Universal Robots PolyScope program: Sub_Action_V2.urp

Program Sub_Action_V2 (installation=uLM011 MiR C1 BioRad directory=/programs/03 Sub Routines createdIn=5.16.0 lastSavedIn=5.16.0 robotSerialNumber=20245590045)
Calibrated DH parameters: a=[0.000135, -0.047884, -0.355309, -0.000204, 0.00003, 0]; d=[0.162633, 288.058298, -225.853183, -62.071663, 0.099761, 0.099601]; alpha=[1.569987, -0.001468, 0.002675, 1.570079, -1.570235, 0]; deltaTheta=[0, -1.458004, 8.179183, -0.437996, 0.000001, 0]
InitVariablesNode variables(variable(name=CMD_Abort, expression=False), variable(name=CMD_Clear, expression=False))
BeforeStart
  Script file /programs/04 Scripts/001 SCRIPT Errors and Warnings Deifnes V0.2.script
    | #*****************************************************
    | # customer          :   UK Essen
    | # project name      :   P1132
    | #****************************************************
    | # controller        :
    | # software          :
    | #****************************************************
    | # author            :   E.Petrichenko
    | # Copyright (c)     :   United Robotics Group Health and Food GmbH
    | #                       An der Riede 2
    | #                       28816 Stuhr
    | #                       Germany
    | #****************************************************
    | # description       :   centrifuge actions for the application
    | # version:      	:   0.1
    | # created           :   22.08.2024
    | # updated           :
    | #****************************************************
    | # modifications     :
    | #
    | # date              :
    | # name              :
    | # reason            :
    | #****************************************************
    | 
    | 
    | #################################### VARIABLES DEFINITIONS ###################################
    | 
    | ERROR_POSE_NOT_REACHABLE = 1002
    | ERROR_ROBOT_ARM_NOT_IN_HOME_POSE = 1006
    | ERROR_NO_OBJECT_TO_PICK = 1010
    | ERROR_NOT_DOCKED = 2003
    | ERROR_NOT_REACHABLE_TARGET = 2007
    | ERROR_CHARGING_NOT_STARTED = 2008
    | ERROR_AMR_WRONG_MODE = 2009
    | ERROR_UNKNOWN_POSE = 2010
    | ERROR_NO_LANDMARK = 3002
    | ERROR_WRONG_ORDER = 4002
    | ERROR_CENTRIFUGE_CONNECTION = 5001
    | ERROR_CENTRIFUGE_POWER = 5002
    | ERROR_CENTRIFUGE = 5003
    | ERROR_CENTRIFUGE_LID = 5004
    | ERROR_CANNOT_OPEN_HATCH = 5006
    | ERROR_CANNOT_CLOSE_HATCH = 5008
    | ERROR_CANNOT_ROTATE = 5010
    | ERROR_CANNOT_START = 5011
    | ERROR_WRONG_KEY_POSE = 5012
    | ERROR_MISSIING_CENTRACK = 5013
    | 
    | WARNING_POSE_NOT_REACHABLE = 1002
    | WARNING_BATTERY_LEVEL = 2002
    | WARNING_NOT_REACHABLE_TARGET = 2007
    | 
    | 
    | ERROR = struct(
    |     FLAG = False,
    |     ID = 0,
    |     MSG = "")
    | 
    | WARNING = struct(
    |     FLAG = False,
    |     ID = 0,
    |     MSG = "")
    | 
    | 
    | #################################### FUNCTIONS ###################################
    | 
    | def set_error(error_id):
    |     ERROR.ID = error_id
    |     if (ERROR.ID == 0):
    |         ERROR.FLAG = False
    |         ERROR.MSG = ""
    |     else:
    |         ERROR.FLAG = True
    |         if(ERROR.ID == ERROR_POSE_NOT_REACHABLE):
    |             ERROR.MSG = "Pose is not reachable"
    |         elif(ERROR.ID == ERROR_NO_OBJECT_TO_PICK):
    |             ERROR.MSG = "No object to pick"
    |         elif(ERROR.ID == ERROR_NO_LANDMARK):
    |             ERROR.MSG = "No landmark detected"
    |         elif(ERROR.ID == ERROR_ROBOT_ARM_NOT_IN_HOME_POSE):
    |             ERROR.MSG = "Robot arm cannot go to home pose"
    |         elif(ERROR.ID == ERROR_AMR_WRONG_MODE):
    |             ERROR.MSG = "AMR is in the wrong mode"
    |         elif(ERROR.ID == ERROR_NOT_DOCKED):
    |             ERROR.MSG = "Could not dock to the charger"
    |         elif(ERROR.ID == ERROR_NOT_REACHABLE_TARGET):
    |             ERROR.MSG = "Could not reach the target"
    |         elif(ERROR.ID == ERROR_CHARGING_NOT_STARTED):
    |             ERROR.MSG = "Could not start charging"
    |         elif(ERROR.ID == ERROR_UNKNOWN_POSE):
    |             ERROR.MSG = "Unknown navigation target"
    |         elif(ERROR.ID == ERROR_CANNOT_OPEN_HATCH):
    |             ERROR.MSG = "Centrifuge Cannot open the hatch"
    |         elif(ERROR.ID == ERROR_CENTRIFUGE_CONNECTION):
    |             ERROR.MSG = "Cannot reach centrifuge"
    |         elif (ERROR.ID == ERROR_CANNOT_CLOSE_HATCH):
    |             ERROR.MSG = "Centrifuge Cannot close the hatch"
    |         elif (ERROR.ID == ERROR_CANNOT_START):
    |             ERROR.MSG = "Centrifuge Cannot start"
    |         elif (ERROR.ID == ERROR_CANNOT_ROTATE):
    |             ERROR.MSG = "Centrifuge Cannot rotate the rotor"
    |         elif (ERROR.ID == ERROR_WRONG_ORDER):
    |             ERROR.MSG = "Wrong parameter was recieved"
    |         elif (ERROR.ID == ERROR_CENTRIFUGE):
    |             ERROR.MSG = "Centrifuge is in Error"
    |         elif (ERROR.ID == ERROR_WRONG_KEY_POSE):
    |             ERROR.MSG = "Key is in the wrong position"
    |         elif(ERROR.ID == ERROR_MISSIING_CENTRACK):
    |             ERROR.MSG = "Missing rack for centrifuge set"
    |         elif(ERROR.ID == ERROR_CENTRIFUGE_POWER):
    |             ERROR.MSG = "Centrifuge is turned off"
    |         elif(ERROR.ID == ERROR_CENTRIFUGE_LID):
    |             ERROR.MSG = "Lid of the centrifuge is opened"
    |         else:
    |             ERROR.MSG = "Unknown code"
    |         end
    |         textmsg("ERROR:",ERROR)
    |     end
    | end
    | 
    | def set_warning(warning_id):
    |     WARNING.ID = warning_id
    |     if (WARNING.ID == 0):
    |         WARNING.FLAG = False
    |         WARNING.MSG = ""
    |     else:
    |         WARNING.FLAG = True
    |         if(WARNING.ID == WARNING_POSE_NOT_REACHABLE):
    |             WARNING.MSG = "Pose is not reachable"
    |         elif(WARNING.ID == WARNING_BATTERY_LEVEL):
    |             WARNING.MSG = "Batery level dropped to a certain level"
    |         elif(WARNING.ID == WARNING_NOT_REACHABLE_TARGET):
    |             WARNING.MSG = "Not reachable location of AMR"
    |         else:
    |             WARNING.MSG = "Unknown code"
    |         end
    |         textmsg("WARNING:",WARNING)
    |     end
    | end
    | 
    | 
    | def reset_error():
    |   ERROR.ID = 0
    |   ERROR.FLAG = False
    |   ERROR.MSG = ""
    | end
    | 
    | 
    | def reset_warning():
    |     WARNING.ID = 0
    |     WARNING.FLAG = False
    |     WARNING.MSG = ""
    |   end
  Script file /programs/04 Scripts/SCRIPT Transitions V5.2.script
    | #*****************************************************
    | # customer          :   INTERNAL
    | # project name      :
    | #****************************************************
    | # controller        :   UR
    | # software          :   5.13
    | #****************************************************
    | # author            :   P. Koehnke
    | # Copyright (c)     :   United Robotics Group
    | #                       An der Riede 2
    | #                       28816 Stuhr
    | #                       Germany
    | #****************************************************
    | # description       :   transition between workareas
    | # version:      	:   1.2
    | # created           :   28.02.2024
    | # updated           :
    | #****************************************************
    | # modifications     :
    | #
    | # date              :
    | # name              :
    | # reason            :
    | #****************************************************
    | 
    | ######################### further development #########################
    | #   - that the robot can switch the configuration, if necessary
    | #   - introduction of structs
    | #######################################################################
    | 
    | ######################### to be adjusted #########################
    | local WORKAREA_1 = [-0.290,-0.560,-0.001, 0.290, 0.100, 1.000]    # workarea 1 (platform)
    | local WORKAREA_2 = [-1.000,-1.000,-1.000,-0.290, 0.100, 1.000]    # workarea 2 (front right)
    | local WORKAREA_3 = [-1.000, 0.100,-1.000, 0.000, 1.000, 1.000]    # workarea 3 (back right)
    | local WORKAREA_4 = [ 0.000, 0.100,-1.000, 1.000, 1.000, 1.000]    # workarea 4 (back left)
    | local WORKAREA_5 = [ 0.290,-1.000,-1.000, 1.000, 0.100, 1.000]    # workarea 5 (front left)
    | local WORKAREA_6 = [-0.290,-1.000,-1.000, 0.290,-0.560, 1.000]    # workarea 6 (front front)
    | local WORKAREA_7 = [0,0,0,0,0,0]    # reserved
    | local WORKAREA_8 = [0,0,0,0,0,0]    # reserved
    | local WORKAREA_9 = [0,0,0,0,0,0]    # reserved
    | local WORKAREA_10 = [0,0,0,0,0,0]   # reserved
    | 
    | local PSE_WA_1 = p[ 0.000,-0.400, 0.300, 0.000, 0.000, 0.000]
    | local PSE_WA_2 = p[-0.300,-0.300, 0.300, 0.000, 0.000, d2r(-90)]
    | local PSE_WA_3 = p[-0.300, 0.300, 0.300, 0.000, 0.000, d2r(-135)]
    | local PSE_WA_4 = p[ 0.300, 0.300, 0.300, 0.000, 0.000, d2r(135)]
    | local PSE_WA_5 = p[ 0.300,-0.300, 0.300, 0.000, 0.000, d2r(90)]
    | local PSE_WA_6 = p[ 0.000,-0.600, 0.300, 0.000, 0.000, 0.000]       # reserved
    | local PSE_WA_7 = p[ 0.000, 0.000, 0.000, 0.000, 0.000, 0.000]       # reserved
    | local PSE_WA_8 = p[ 0.000, 0.000, 0.000, 0.000, 0.000, 0.000]       # reserved
    | local PSE_WA_9 = p[ 0.000, 0.000, 0.000, 0.000, 0.000, 0.000]       # reserved
    | local PSE_WA_10 = p[ 0.000, 0.000, 0.000, 0.000, 0.000, 0.000]      # reserved
    | 
    | local JNT_STANDARD_C1 = [ 1.57,-1.57, 1.57,-1.57,-1.57,0]
    | local JNT_STANDARD_C2 = [-1.57,-1.57,-1.57,-1.57, 1.57,0]
    | local CLEARANCE_STANDARD = [-0.500,-0.900,-1.000, 0.500, 0.900, 1.000]  # desired free space around the base
    | local DISTANCE_TO_CLEARANCE = 0.300
    | local RADIUS_HELPER_POSES = 0.250
    | local RADIUS_TRANSITION_POSES = 0.400
    | local workareas = [WORKAREA_1, WORKAREA_2, WORKAREA_3, WORKAREA_4, WORKAREA_5, WORKAREA_6, WORKAREA_7, WORKAREA_8, WORKAREA_9, WORKAREA_10]
    | local poses = [PSE_WA_1, PSE_WA_2, PSE_WA_3, PSE_WA_4, PSE_WA_5, PSE_WA_6, PSE_WA_7, PSE_WA_8, PSE_WA_9, PSE_WA_10]
    | 
    | ######################### end of adjustment #########################
    | 
    | local pi = 3.14159265
    | local axis_config_current = 0
    | local axis_config_new = 0
    | local workarea_current = 0
    | local workarea_new = 0
    | local reverse_rotation = False
    | local yaw_locked =  0
    | local pose_start = struct(crt = p[0,0,0,0,0,0], jnt = [0,0,0,0,0,0], q = [0,0,0,0,0,0])
    | local pose_help = struct(crt = p[0,0,0,0,0,0], jnt = [0,0,0,0,0,0], q = [0,0,0,0,0,0])
    | local pose_target = struct(crt = p[0,0,0,0,0,0], jnt = [0,0,0,0,0,0], q = [0,0,0,0,0,0])
    | local pose = struct(crt = p[0,0,0,0,0,0], jnt = [0,0,0,0,0,0], q = [0,0,0,0,0,0])
    | 
    | def get_tool_free_pose(pose_ref=get_actual_tcp_pose(), dir=[0,0,0], move_in_base_frame=False):
    |     # get a recovery pose
    |     # dir is providing the direction and distance in X, Y and Z
    |     # if 'move_in_base_frame' is set, dir will be interpreted as absolute values for a movement in base frame
    | 
    |     local pose_target = pose_ref
    |     local i = 0
    | 
    |     if (move_in_base_frame):
    |         while (i<3):
    |             # move only,
    |             # if the demanded position is bigger than zero and the current position is below the demanded one or
    |             # if the demanded position is smaller than zero and the current position is above the demanded one
    |             if ((dir[i]>0 and pose_ref[i]<dir[i]) or (dir[i]<0 and pose_ref[i]>dir[i])):
    |                 pose_target[i] = dir[i]
    |             end
    |             i = i + 1
    |         end
    |     else:
    |         pose_target = pose_trans(pose_ref, p[dir[0], dir[1], dir[2], 0, 0, 0])
    |     end
    | 
    |     return pose_target
    | end
    | 
    | def check_workarea(reference_pose):
    |     # the actual TCP position is compared to predefined areas (cubic) to determine in which area the robot arm is
    |     # a workarea is defined as a list of coordinates, where the first 3 values are X, Y, and Z with the smallest values and
    |     # the next 3 values specify X, Y and Z for the biggest values
    | 
    |     local data_size = size(workareas)
    |     local i = 0
    |     local size_workarea = p[0,0,0,0,0,0]
    |     local pose_workarea = p[0,0,0,0,0,0]
    | 
    |     while (i < data_size[0]):
    |         pose_workarea = pose_trans(inv(p[workareas[i, 0], workareas[i, 1], workareas[i, 2], 0, 0, 0]), reference_pose)
    |         size_workarea = pose_sub(p[workareas[i, 3], workareas[i, 4], workareas[i, 5], 0, 0, 0], p[workareas[i, 0], workareas[i, 1], workareas[i, 2], 0, 0, 0])
    |         if  ((pose_workarea[0]>0 and pose_workarea[0]<size_workarea[0]) and
    |             (pose_workarea[1]>0 and pose_workarea[1]<size_workarea[1]) and
    |             (pose_workarea[2]>0 and pose_workarea[2]<size_workarea[2])):
    |             return i + 1
    |         end
    |         i = i + 1
    |     end
    |     return 0
    | end
    | 
    | def check_current_axis_config():
    |     # function determnines, if the arm is oriented in one or the other configuration.
    |     # it means, that the ellbow joint is flipped and so are the wrist joints.
    | 
    |     local jnt_current = get_actual_joint_positions()
    | 
    |     # ellbow has positiv angle
    |     if (jnt_current[2]> 0):
    |         return 1
    |     # ellbow has negativ angle
    |     elif (jnt_current[2]< 0):
    |         return 2
    |     # angle is 0
    |     else:
    |         return 0
    |     end
    | end
    | 
    | def switch_axis_config(axis_config):
    |     # function to switch betwwen the axis configuration 1 and 2.
    | 
    |     if (axis_config == 1):
    |         return 2
    |     elif (axis_config ==2):
    |         return 1
    |     end
    | end
    | 
    | def get_transition_pose(workarea, axis_config, closest=False, keep_xyz=[False, False, False]):
    |     # get the correspondig pose from the list of poses
    | 
    |     local jnt_current = get_actual_joint_positions()
    |     local pose_current = get_actual_tcp_pose()
    |     local i = 0
    | 
    |     pose.crt = poses[workarea-1]
    |     # if wanted, the pose will take the current position as desired x, y and z
    |     while (i < 3):
    |         if keep_xyz[i]:
    |             pose.crt[i] = pose_current[i]
    |         end
    |         i = i + 1
    |     end
    | 
    |     if (axis_config == 1):
    |         pose.q = JNT_STANDARD_C1
    |     elif (axis_config == 2):
    |         pose.q = JNT_STANDARD_C2
    |     end
    | 
    |     if closest:
    |         pose.q[0] = jnt_current[0]
    |     end
    | 
    |     if get_inverse_kin_has_solution(pose.crt, qnear=pose.q):
    |         pose.jnt = get_inverse_kin(pose.crt, qnear=pose.q)
    |     else:
    |         popup("no solution found for the transition pose", blocking= True)
    |     end
    | 
    |     return pose
    | end
    | 
    | def get_transition_pose_2(ref, radius, axis_config, closest=False):
    |     # get the correspondig pose from the list of poses
    | 
    |     local jnt_current = get_actual_joint_positions()
    |     local yaw_current = get_yaw_too_base(ref)
    | 
    |     #pose.crt = get_tool_free_pose(pose_ref=ref, dir=[0, 0, DISTANCE_TO_CLEARANCE], move_in_base_frame=True)
    | 
    |     if (axis_config == 1):
    |         pose.q = JNT_STANDARD_C1
    |     elif (axis_config == 2):
    |         pose.q = JNT_STANDARD_C2
    |     end
    | 
    |     if closest:
    |         pose.q[0] = jnt_current[0]
    |     end
    | 
    |     # get coordinates of the circle with the same angle as the given pose to the
    |     if ref == p[0,0,0,0,0,0]:
    |         pose.crt = PSE_WA_1
    |     else:
    |         pose.crt =
    |         p[radius * cos(yaw_current-pi/2),
    |         radius * sin(yaw_current-pi/2),
    |         DISTANCE_TO_CLEARANCE,
    |         0,
    |         0,
    |         yaw_current + get_locked_yaw()]
    |     end
    | 
    |     if get_inverse_kin_has_solution(pose.crt, qnear=pose.q):
    |         pose.jnt = get_inverse_kin(pose.crt, qnear=pose.q)
    |         #return pose
    |     else:
    |         popup("no solution found for the transition pose", blocking= True)
    |     end
    | 
    |     return pose
    | end
    | 
    | def get_rounded_mm(value):
    |     if (value < 0):
    |         return ceil(value*1000)
    |     elif (value >= 0):
    |         return floor(value*1000)
    |     end
    | end
    | 
    | def get_yaw_too_base(pose):
    |     # get the yaw relative to the base frame
    |     local pose_x_mm = 0
    |     local pose_y_mm = 0
    |     local yaw = 0
    | 
    |     pose_x_mm = get_rounded_mm(pose[0])
    |     pose_y_mm = get_rounded_mm(pose[1])
    | 
    |     if (pose_x_mm == 0 and pose_y_mm < 0):
    |         yaw = 0
    |     elif (pose_x_mm == 0 and pose_y_mm > 0):
    |         yaw = pi
    |     elif (pose_x_mm < 0 and pose_y_mm == 0):
    |         yaw = -pi/2
    |     elif (pose_x_mm > 0 and pose_y_mm == 0):
    |         yaw = pi/2
    |     else:
    |         yaw = atan2(pose[0], pose[1])
    |         if (-pi < yaw) and (yaw < 0):
    |             yaw = - yaw - pi
    |         elif (0 < yaw) and (yaw < pi):
    |             yaw = - yaw + pi
    |         else:
    |             yaw = pi
    |         end
    |     end
    |     return yaw
    | end
    | 
    | def get_helper_pose():
    |     # get the helper pose, as described
    | 
    |     local m_line = 0                    # slope of the line between base and circle point
    |     local n = 0                         # shift on the ordinate axis
    |     local m_normal = 0                  # slope of the normal of the line between base and circle point
    |     local x_p1 = 0                      # x coordinate of first circle point
    |     local x_p2 = 0                      # x coordinate of second circle point
    |     local y_p1 = 0                      # y coordinate of first circle point
    |     local y_p2 = 0                      # y coordinate of second circle point
    |     local jnt_help_1 = [0,0,0,0,0,0]
    |     local jnt_help_2 = [0,0,0,0,0,0]
    | 
    |     if (pose_start.crt != pose_target.crt):
    |         if (pose_start.crt[0] == pose_target.crt[0]):
    |             m_normal = 0
    |         elif (pose_start.crt[0] != pose_target.crt[0]):
    |             m_line = (pose_target.crt[1]-pose_start.crt[1])/(pose_target.crt[0]-pose_start.crt[0])    # calculation of the slope between start and target
    |             n = pose_start.crt[1] - m_line * pose_start.crt[0]
    |         end
    |         if (-0.00001 > m_line or m_line > 0.00001):
    |             m_normal = -1/m_line
    |         end
    | 
    |         # using p-q-formula for getting the crossing points
    |         x_p1 = sqrt(pow(RADIUS_HELPER_POSES, 2)/(pow(m_normal, 2)+1)) * -1
    |         x_p2 = sqrt(pow(RADIUS_HELPER_POSES, 2)/(pow(m_normal, 2)+1))
    |         y_p1 = m_normal * x_p1
    |         y_p2 = m_normal * x_p2
    |         pose.q = pose_start.jnt
    | 
    |         if (point_dist(pose_start.crt, p[x_p1, y_p1,0,0,0,0]) < point_dist(pose_start.crt, p[x_p2, y_p2,0,0,0,0])):
    |             if reverse_rotation:
    |                 pose_help.crt[0] = x_p2
    |                 pose_help.crt[1] = y_p2
    |                 pose.q = pose_target.jnt
    |             else:
    |                 pose_help.crt[0] = x_p1
    |                 pose_help.crt[1] = y_p1
    |                 pose.q = pose_start.jnt
    |             end
    |         elif (point_dist(pose_start.crt, p[x_p1, y_p1,0,0,0,0]) > point_dist(pose_start.crt, p[x_p2, y_p2,0,0,0,0])):
    |             if reverse_rotation:
    |                 pose_help.crt[0] = x_p1
    |                 pose_help.crt[1] = y_p1
    |                 pose.q = pose_target.jnt
    |             else:
    |                 pose_help.crt[0] = x_p2
    |                 pose_help.crt[1] = y_p2
    |                 pose.q = pose_start.jnt
    |             end
    |         elif (point_dist(pose_start.crt, p[x_p1, y_p1,0,0,0,0]) == point_dist(pose_start.crt, p[x_p2, y_p2,0,0,0,0])):
    |             jnt_help_1 = get_inverse_kin(p[x_p1, y_p1,pose_start.crt[2],pose_start.crt[3],pose_start.crt[4],pose_start.crt[5]], qnear=pose.q)
    |             jnt_help_2 = get_inverse_kin(p[x_p2, y_p2,pose_start.crt[2],pose_start.crt[3],pose_start.crt[4],pose_start.crt[5]], qnear=pose.q)
    |             if (pose_start.jnt[0]<jnt_help_1[0] and jnt_help_1[0]<pose_target.jnt[0]) or (pose_start.jnt[0]>jnt_help_1[0] and jnt_help_1[0]>pose_target.jnt[0]):
    |                 pose_help.crt[0] = x_p1
    |                 pose_help.crt[1] = y_p1
    |             elif (pose_start.jnt[0]<jnt_help_2[0] and jnt_help_2[0]<pose_target.jnt[0]) or (pose_start.jnt[0]>jnt_help_2[0] and jnt_help_2[0]>pose_target.jnt[0]):
    |                 pose_help.crt[0] = x_p2
    |                 pose_help.crt[1] = y_p2
    |             end
    |             pose.q = pose_start.jnt
    |         end
    | 
    |         pose_help.crt[2] = 0.5 * (pose_start.crt[2] + pose_target.crt[2])
    | 
    |         if ((pose_start.crt[1] < 0 and pose_target.crt[1] > 0) or (pose_start.crt[1] > 0 and pose_target.crt[1] < 0)):
    |             if get_inverse_kin_has_solution(pose.crt, qnear=pose.q):
    |                 pose.jnt = get_inverse_kin(pose.crt, qnear=pose.q)
    |             else:
    |                 popup("no solution found for the helper pose", blocking= True)
    |             end
    |         end
    |     end
    |     return pose
    | end
    | 
    | def adjust_transition_poses(pose_identifier):
    |     # adjust the orientation of the transition poses by determining the the current orientation
    | 
    |     local pose_current = get_actual_tcp_pose()
    |     local jnt_current = get_actual_joint_positions()
    |     local rpy_current = rotvec2rpy([pose_current[3],pose_current[4],pose_current[5]])
    |     local rotvec_new = [0,0,0]
    | 
    |     if (pose_identifier == "start"):
    |         pose.q = pose_start.jnt
    |         pose.crt = get_forward_kin(pose_start.jnt)
    |     elif (pose_identifier == "helper"):
    |         pose.q = pose_help.jnt
    |         pose.crt = get_forward_kin(pose_help.jnt)
    |     elif (pose_identifier == "target"):
    |         pose.q = pose_target.jnt
    |         pose.crt = get_forward_kin(pose_target.jnt)
    |     end
    | 
    |     rotvec_new = rpy2rotvec([rpy_current[0], rpy_current[1], get_yaw_too_base(pose.crt) + yaw_locked])
    |     pose.crt = p[pose.crt[0], pose.crt[1], pose.crt[2], rotvec_new[0], rotvec_new[1], rotvec_new[2]]
    | 
    |     pose.q[3] = jnt_current[3]
    |     pose.q[4] = jnt_current[4]
    |     pose.q[5] = jnt_current[5]
    |     if get_inverse_kin_has_solution(pose.crt, qnear=pose.q) and is_within_safety_limits(pose.crt):
    |         pose.jnt = get_inverse_kin(pose.crt, qnear=pose.q)
    |     else:
    |         popup(str_cat("no solution for ", pose_identifier), error=True, blocking=True)
    |     end
    |     return pose.jnt
    | end
    | 
    | def get_locked_yaw():
    |     local pose_current = get_actual_tcp_pose()
    |     local rpy_current = rotvec2rpy([pose_current[3],pose_current[4],pose_current[5]])
    |     local rotvec_new = rpy2rotvec([rpy_current[0], rpy_current[1], get_yaw_too_base(pose_current)])
    |     local pose_reference = p[pose_current[0], pose_current[1], pose_current[2], rotvec_new[0], rotvec_new[1], rotvec_new[2]]
    |     local pose_to_reference = pose_trans(pose_inv(pose_reference), get_actual_tcp_pose())
    |     yaw_locked = pose_to_reference[5]
    | 
    |     return yaw_locked
    | end
    | 
    | def do_transition(reference_pose=p[0,0,0,0,0,0], mode=2, keep_xyz=[False, False, False], keep_rxry=False, a=1.4, v=1.05, r=0.100):
    |     # the robot will evaluate the current and target workarea
    |     # after that, the robot will move between the workareas automatically.
    |     # parameters:
    |     # reference_pose:   a pose/frame were the robot should work next. If nothing is given, base frame will be used as target
    |     # keep_rxry:        if true, the robot will keep the orientation of the tool during the movement
    | 
    |     ################# checking #################
    |     axis_config_current = check_current_axis_config()           # 0: unknown, 1: config 1, 2: config 2
    |     workarea_current = check_workarea(get_actual_tcp_pose())    # between 0 and the amount of defined workareas
    |     workarea_new = check_workarea(reference_pose)               # between 0 and the amount of defined workareas
    |     if(workarea_current==workarea_new):
    |          return 0
    |     end
    |     if (workarea_current != 0 and workarea_new != 0):
    |         ################# get axisvalues #################
    |         # pose_start = get_transition_pose(workarea_current, axis_config_current, closest=not reverse_rotation, keep_xyz=keep_xyz)
    |         pose_start = get_transition_pose_2(get_actual_tcp_pose(), RADIUS_TRANSITION_POSES, axis_config_current, closest=not reverse_rotation)
    |         if (workarea_current == 3 and workarea_new == 4) or (workarea_current == 4 and workarea_new == 3):
    |             # pose_target = get_transition_pose(workarea_new, axis_config_current, closest=True)
    |             pose_target = get_transition_pose_2(reference_pose, RADIUS_TRANSITION_POSES, axis_config_current, closest=True)
    |             reverse_rotation = True
    |         else:
    |             pose_target = get_transition_pose_2(reference_pose, RADIUS_TRANSITION_POSES, axis_config_current, closest=(workarea_current == workarea_new))
    |             if reverse_rotation:
    |                 reverse_rotation = False
    |             end
    |         end
    |         # pose_help = get_helper_pose()
    |         global A_Start = pose_start.crt
    |         global A_Help = pose_help.crt
    |         global A_End = pose_target.crt
    | 
    | 
    |         ################# adjustments #################
    |         if (keep_rxry):
    |             get_locked_yaw()
    |             if (pose_start.jnt == pose_target.jnt):
    |                 pose_target.jnt = adjust_transition_poses("target")
    |                 pose_start.jnt = pose_target.jnt
    |             else:
    |                 pose_start.jnt = adjust_transition_poses("start")
    |                 pose_target.jnt = adjust_transition_poses("target")
    |             end
    |             if (pose_help.jnt != [0,0,0,0,0,0]):
    |                 pose_help.jnt = adjust_transition_poses("helper")
    |             end
    |         end
    | 
    |         global A_Start = pose_start.crt
    |         global A_Help = pose_help.crt
    |         global A_End = pose_target.crt
    | 
    |         ################# movements #################
    | 
    |         if point_dist(pose_start.crt, pose_target.crt) > 0.100:
    |             movej(pose_start.jnt, a=a, v=v, r=r)
    |         end
    |         # if (pose_help.jnt != [0,0,0,0,0,0]):
    |         #     movej(pose_help.jnt, a=a, v=v, r=r)
    |         # end
    |         movej(pose_target.jnt, a=a, v=v)
    |     else:
    |         # define error
    |     end
    | 
    |     ################# checking #################
    |     axis_config_current = check_current_axis_config()           # 0: unknown, 1: config 1, 2: config 2
    |     workarea_current = check_workarea(get_actual_tcp_pose())    # between 0 and the amount of defined workareas
    | end
  Script file /programs/04 Scripts/SCRIPT Utility V5.1.script
    | #*****************************************************
    | # customer          :   tbd
    | # project name      :   tbd
    | #****************************************************
    | # controller        :
    | # software          :
    | #****************************************************
    | # author            :   P. Koehnke (+49 1628859904; p.koehnke@unitedrobotics.group)
    | # Copyright (c)     :   United Robotics Group Health and Food GmbH
    | #                       An der Riede 2
    | #                       28816 Stuhr
    | #                       Germany
    | #****************************************************
    | # description       :   utility programs for the application
    | # version:      	:   3.1
    | # created           :   30.01.2023
    | # updated           :
    | #****************************************************
    | # modifications     :   get_tool_free_pose_2(), get_index_from_list()
    | #
    | # date              :   05.01.2024
    | # name              :   PK
    | # reason            :
    | #****************************************************
    | 
    | def found_in_matrix(data, req_id, req_idx):
    |     local id = -1
    |     local dimensions = size(data)
    |     local loop_dataset = 0
    | 
    |     while (id != req_id and loop_dataset < dimensions[0]):
    |         id = data[loop_dataset, 0]
    |         if (id == req_id):
    |             return data[loop_dataset, req_idx]
    |         else:
    |             loop_dataset = loop_dataset + 1
    |         end
    |     end
    | end
    | 
    | def found_in_list(value, list):
    |     local idx = 0
    | 
    |     while (idx < length(list)):
    |         if (value == list[idx]):
    |             return True
    |         end
    |         idx = idx + 1
    |     end
    |     return False
    | end
    | 
    | def get_index_from_list(list, value=-1):
    |     local idx = 0
    | 
    |     while (idx < length(list)):
    |         if (value == -1):
    |             if (list[idx] != 0):
    |                 return idx
    |             end
    |         else:
    |             if (list[idx] == value):
    |                 return idx
    |             end
    |         end
    |         idx = idx + 1
    |     end
    |     return -1
    | end
    | 
    | def pose_RPY2RotVec(pose):
    |     local rotvec = rpy2rotvec([d2r(pose[3]),d2r(pose[4]),d2r(pose[5])])
    |     return p[pose[0],pose[1],pose[2],rotvec[0],rotvec[1],rotvec[2]]
    | end
    | 
    | def pose_RotVec2RPY(pose):
    |     local rpy = rotvec2rpy([pose[3],pose[4],pose[5]])
    |     return p[pose[0],pose[1],pose[2],r2d(rpy[0]),r2d(rpy[1]),r2d(rpy[2])]
    | end
    | 
    | def swivel(frame_ref, angles=[0,0,0], pose=p[0,0,0,0,0,0]):
    | 
    |     local rpy_ref = [0,0,0]
    |     local rpy_new = [0,0,0]
    |     local rotvec_new = [0,0,0]
    |     local pose_from = p[0,0,0,0,0,0]
    |     local pose_to = p[0,0,0,0,0,0]
    |     local i = 0
    | 
    |     if (pose == p[0,0,0,0,0,0]):
    |         pose_to = pose_trans(pose_inv(frame_ref), get_actual_tcp_pose())
    |     else:
    |         pose_to = pose
    |     end
    | 
    |     rpy_ref = rotvec2rpy(frame_ref[3], frame_ref[4], frame_ref[5])
    | 
    |     while (i < 3):
    |         rpy_new[i] = rpy_ref[i] + d2r(angles[i])
    |         i = i + 1
    |     end
    | 
    |     rotvec_new = rpy2rotvec(rpy_new)
    |     pose_from = p[0,0,0,rotvec_new[0],rotvec_new[1],rotvec_new[2]]
    |     pose_to = p[pose_to[0], pose_to[1], pose_to[2], rotvec_new[0], rotvec_new[1], rotvec_new[2]]
    | 
    |     return pose_trans(pose_from, pose_to)
    | end
    | 
    | def get_random_pose(pose_ref, mode="", range_max=[0,0,0]):
    |     # modi: "cubic", "rotation"
    |     # getting a random pose in the x/y-plane. range can be set for each
    |     # translation and rotation.
    |     local rpy_random = [0,0,0]
    |     local rotvec_random = [0,0,0]
    |     local pose_random = pose_ref
    |     local i = 0
    | 
    |     if (mode == "cubic"):
    |         # cubic mode: random pose takes only x, y and z
    |         i = 0
    |         while(i<3):
    |             pose_random[i] = pose_ref[i] + range_max[i] * (random() - 0.5)
    |             i = i + 1
    |         end
    |         return pose_random
    | 
    |     elif (mode == "rotation"):
    |         i = 0
    |         while(i<3):
    |             rpy_random[i] = d2r(range_max[i]) * (random() - 0.5)
    |             i = i + 1
    |         end
    |         rotvec_random = rpy2rotvec(rpy_random)
    |         pose_random = pose_trans(p[0,0,0,rotvec_random[0],rotvec_random[1],rotvec_random[2]], pose_ref)
    |         return pose_random
    | 
    |     else:
    |         # unknown mode, return pose_ref
    |         return pose_ref
    |     end
    | end
    | 
    | def get_pattern_pos_rectangle(counter, direction, patternsize, patterninc=[0,0], patternwidth=[0,0]):
    |     # defines the position inside a rectangular pattern
    |     # patternsize describes, how many objects are in x-direction and how many in y-direction [x, y]
    |     # patternwidth will give the total length of each direction [x, y]
    |     local X_Fac = 0
    |     local Y_Fac = 0
    |     local max = patternsize[0]*patternsize[1]
    | 
    |     if (1>counter or counter>max):
    |         counter = 1
    |     end
    | 
    |     if (direction == "Y" or direction == "y"):
    |         X_Fac = floor((counter - 1) / patternsize[1])
    |         Y_Fac = (counter - 1) % patternsize[1]
    |     elif (direction == "X" or direction == "x"):
    |         X_Fac = (counter - 1) % patternsize[0]
    |         Y_Fac = floor((counter - 1) / patternsize[0])
    |     end
    | 
    |     if patternwidth != [0,0]:
    |         patterninc = [patternwidth[0]/(patternsize[0]-1), patternwidth[1]/(patternsize[1]-1)]
    |     end
    | 
    |     return p[X_Fac*patterninc[0], Y_Fac*patterninc[1],0,0,0,0]
    | end
    | 
    | def get_pattern_pos_circle(counter, radius, angle, direction, pattern, patternsize=[0,0]):
    |     # get the patternpos for a circular pattern through a counter
    |     # need the radius and the angle in radiants
    |     local X_Fac = 0
    |     local Y_Fac = 0
    |     local rad_bow = 0
    |     local radius_cal = 0
    |     local ref = p[0,0,0,0,0,0]
    | 
    |     if (direction == "Y" or direction == "y"):
    |         X_Fac = floor((counter - 1) / pattern[1])
    |         Y_Fac = (counter - 1) % pattern[1]
    |     elif (direction == "X" or direction == "x"):
    |         X_Fac = (counter - 1) % pattern[0]
    |         Y_Fac = floor((counter - 1) / pattern[0])
    |     end
    | 
    |     # the opening angle will be calculated in x-direction
    |     # works only between -90 and 90 degree
    |     rad_bow = -angle/(pattern[0]-1) * X_Fac + angle/2
    | 
    |     if (counter%2 == 0):
    |         radius_cal = radius - patternsize[1]/(pattern[1])
    |     else:
    |         radius_cal = radius + patternsize[1]/(pattern[1])
    |     end
    |     ref = p[0, radius_cal, 0, 0, 0, 0]
    | 
    |     return p[ref[0]*cos(rad_bow)-ref[1]*sin(rad_bow), (ref[0]*sin(rad_bow)+ref[1]*cos(rad_bow))-radius,0,0,0,0]
    | end
    | 
    | def get_pattern_counter(pose, direction, pattern, patterninc=[0,0], patternsize=[0,0]):
    |     # returns the counter for a pattern from a given cartesian pose
    |     local patternpose = p[pose[0],pose[1],0,0,0,0]
    |     local floatFacX = 0.0
    |     local floatFacY = 0.0
    |     local remainder = 0.0
    |     local FacX = 0
    |     local FacY = 0
    | 
    |     # since the pattern spreads from the origin in positive axis-directions, all negative values
    |     # (which could appear due to a position near an axis) will set to zero
    |     if (pose[0]<0):
    |         patternpose = p[0,pose[1],0,0,0,0]
    |     end
    |     if (pose[1]<0):
    |         patternpose = p[pose[0],0,0,0,0,0]
    |     end
    |     # calculate the factor for each axis
    |     floatFacX = patternpose[0]/(patternsize[0]*(pattern[0]-1))
    |     floatFacY = patternpose[1]/(patternsize[1]*(pattern[1]-1))
    |     # determine the remainder after the comma/point
    |     if (floatFacX>1):
    |         remainder = floatFacX%floor(floatFacX)
    |     else:
    |         remainder = floatFacX
    |     end
    |     if (remainder<0.5):
    |         FacX = floatFacX-remainder
    |     else:
    |         FacX = floatFacX+(1-remainder)
    |     end
    | 
    |     if (floatFacY>1):
    |         remainder = floatFacY%floor(floatFacY)
    |     else:
    |         remainder = floatFacY
    |     end
    |     if (remainder<0.5):
    |         FacY = floatFacY-remainder
    |     else:
    |         FacY = floatFacY+(1-remainder)
    |     end
    |     # calculation of the counter in the desired axis-direction
    |     if (direction=="x" or direction=="X"):
    |         return FacX*pattern[1] + FacY + 1
    |     elif (direction=="y" or direction=="Y"):
    |         return FacY*pattern[0] + FacX + 1
    |     end
    | end
    | 
    | def get_plc_reg(mod_sig_name):
    | 	return integer_to_binary_list(modbus_get_signal_status(mod_sig_name))
    | end
    | 
    | def set_plc_reg(mod_sig_name, mod_sig_list):
    | 	modbus_set_output_register(mod_sig_name,binary_list_to_integer(mod_sig_list),False)
    | end
    | 
    | def check_decapping(offset=0, timeout=5):
    |     # checken, ob der Deckel schon ab ist
    |     local start = get_actual_tcp_pose()
    |     local current_offset = 0
    |     local timecounter = 0
    |     while (current_offset < offset):
    |         current_offset = pose_dist(start, get_actual_tcp_pose())
    |         timecounter = timecounter + 1
    |         if (timecounter*0.5 == timeout):
    |             break
    |         end
    |         sleep(0.5)
    |     end
    |     stopl(0.5)
    | end
    | 
    | def check_capping(torque=0):
    |     # checken, wann der Deckel verschraubt ist
    |     force_mode(get_actual_tcp_pose(), [0,0,1,0,0,0], [0,0,-2.0,0,0,0], 2, [0,0,0.100,0,0,0])
    | end
    | 
    | def is_reachable(frame, poses, offsets=[0,0,0]):
    |     local idx = 0
    |     local pose = p[0,0,0,0,0,0]
    | 
    |     while (idx < length(poses)):
    |         pose = poses[idx]
    |         pose[0] = pose[0] + offsets[0]
    |         pose[1] = pose[1] + offsets[1]
    |         pose[2] = pose[2] + offsets[2]
    | 
    |         if pose != p[0,0,0,0,0,0]:
    |             if (not get_inverse_kin_has_solution(pose_trans(frame, pose))):
    |                 textmsg(str_cat(str_cat("Pose ", to_str(idx + 1)), " is not reachable"))
    |                 return False
    |             end
    |         end
    |         idx = idx + 1
    |     end
    |     return True
    | end
    | 
    | def is_within_limits(frame, poses, offsets=[0,0,0]):
    |     local idx = 0
    |     local pose = p[0,0,0,0,0,0]
    | 
    |     while (idx < length(poses)):
    |         pose = poses[idx]
    |         pose[0] = pose[0] + offsets[0]
    |         pose[1] = pose[1] + offsets[1]
    |         pose[2] = pose[2] + offsets[2]
    | 
    |         if is_reachable(frame=frame, poses=poses, offsets=offsets):
    |             if (not is_within_safety_limits(get_inverse_kin(pose_trans(frame, pose), get_actual_joint_positions()))):
    |                 textmsg(str_cat(str_cat("Pose ", to_str(idx + 1)), "is out of joint limits"))
    |                 return False
    |             else:
    |                 idx = idx + 1
    |             end
    |         else:
    |             return False
    |         end
    |     end
    |     return True
    | end
    | 
    | def action_manipulator_decapping():
    |   zero_ftsensor()
    |   local DCP_Start = get_actual_tcp_pose ()
    |   global DCP_Actual = get_actual_tcp_pose ()
    |   local DCP_Height = 0.021
    |   global ForceCounter = 0
    |   sleep(0.02)
    |   zero_ftsensor()
    |   force_mode(p[0.0, 0.0, 0.0, 0.0, 0.0, 0.0], [0, 0, 1, 0, 0, 0], [0.0, 0.0, 17.0, 0.0, 0.0, 10.0], 2, [0.1, 0.1, 0.02, 0.3490658503988659, 0.3490658503988659, 0.3490658503988659])
    |   thread Thread_while_684():
    |     while (True):
    |       global DCP_Actual = get_actual_tcp_pose ()
    |       sleep(0.2)
    |       global ForceCounter = ForceCounter + 1
    |       if (ForceCounter > 30):
    |         zero_ftsensor()
    |         global ForceCounter = 0
    |       end
    |     end
    |   end
    |   if (DCP_Actual[2] <= DCP_Start[2] + DCP_Height):
    |     global thread_handler_decapping = run Thread_while_684()
    |     while (DCP_Actual[2] <= DCP_Start[2] + DCP_Height):
    |       sync()
    |     end
    |     kill thread_handler_decapping
    |   end
    |   end_force_mode()
    |   stopl(5.0)
    | end
  PRC_Target := 0
  PRC_Target := 1
  Action := 1
  Action := 2
  Action := 7
  ITM_ID := 2
  JIG := 1
  JIG_Slot := 2
Robot Program (runOnlyOnce=true)
  Folder PreSettings
    Folder init poses
      PSE_A := p[0,0,0,0,0,0]
      PSE_A_H := p[0,0,0,0,0,0]
      PSE_T := p[0,0,0,0,0,0]
      PSE_T_H := p[0,0,0,0,0,0]
      PSE_G := p[0,0,0,0,0,0]
      PSE_G_H := p[0,0,0,0,0,0]
      PSE_R := p[0,0,0,0,0,0]
      PSE_R_H := p[0,0,0,0,0,0]
      JNT_A := [0,0,0,0,0,0]
      JNT_S := [0,0,0,0,0,0]
      JNT_Q := [0,0,0,0,0,0]
    PROCESS_Info := "work at target, Table"
    PRM_TubHghtDiff := -0.024
    Folder Gripping parameters
      GRP_Open_Pos := 45
      GRP_Close_Pos := 100
      Script: rq_set_force_norm(20)
      Script: rq_set_speed_norm(80)
    Switch expression=ITM_ID
      Case (caseValue=1)
        Folder uML
          Switch expression=JIG
            Case (caseValue=2)
              Folder biorad rack tubes
                GRP_Open_Pos := 60
                FRM_Reference := uLM_BradRckTubs
                Tubes_in_Rack := 6
                PSE_T := pose_RPY2RotVec(p[0.02*(JIG_Slot%Tubes_in_Rack),-0.04365*floor(JIG_Slot/Tubes_in_Rack),0.003,0,0,-90])
                SuppressedNode
                  Script: PSE_T[2]=PSE_T[2]+PRM_TubHghtDiff
                If (JIG_Slot%Tubes_in_Rack)>1
                  Script: PSE_T[0]=PSE_T[0]+0.0165
                  If (JIG_Slot%Tubes_in_Rack)>4
                    Script: PSE_T[0]=PSE_T[0]+0.0235
                    SuppressedNode
                      If (JIG_Slot%10)>6
                        Script: PSE_T[0]=PSE_T[0]+0.0165
                PSE_R := pose_add(PSE_T, p[0,0,0.2500,0,0,0])
                PSE_A := pose_add(PSE_T, p[0,0,0.1,0,0,0])
            Case (caseValue=4)
              Folder centrifuge rack tubes
                GRP_Open_Pos := 60
                FRM_Reference := uLM_CentTubes
                PSE_T := pose_RPY2RotVec(p[0.0975*(JIG_Slot%4),0,0.002,0,0,0])
                SuppressedNode
                  Script: PSE_T[2]=PSE_T[2]+PRM_TubHghtDiff
                If JIG_Slot>3 and JIG_Slot≤7
                  Script: PSE_T[1]=0.06
                  Script: PSE_T[0]=PSE_T[0]+0.06
                ElseIf JIG_Slot>7 and JIG_Slot≤11
                  Script: PSE_T[0]=PSE_T[0]+0.06
                ElseIf JIG_Slot>11 and JIG_Slot≤15
                  Script: PSE_T[1]=0.06
                PSE_R := pose_add(PSE_T, p[0,0,0.150,0,0,0])
                PSE_A := pose_add(PSE_T, p[0,0,0.15,0,0,0])
                JNT_Q := [-1.4,-1.89,-1.4,-1.42,1.57,0.18]
            Case (caseValue=5)
              Folder 3finger gripper
                Folder define poses
                  'Place in 3finger'
                  Script: FRM_Reference = uML_3fingergrip
                  PSE_T := pose_RPY2RotVec(p[0,0,0.003,0,0,0])
                  Script: PSE_T[2]=PSE_T[2]+PRM_TubHghtDiff
                  If Action≟5
                    PSE_T := pose_RPY2RotVec(p[0,0,0.018,0,0,0])
                    PSE_T_H := pose_trans(PSE_T, p[0,0,0.02,0,0,0])
                  If Action≟3
                    Script: PSE_T[5]=PSE_T[5]+d2r(155)
                  PSE_A := pose_trans(PSE_T, p[0,0,0.1,0,0,0])
                  PSE_R := pose_add(PSE_T, p[0,0,0.060,0,0,0])
            Case (caseValue=6)
              Folder Caps bin
                Folder define poses
                  'Drop cap'
                  Script: FRM_Reference=uML_CapBin
                  SuppressedNode
                    PSE_T := pose_RPY2RotVec(p[0.037,0,0.005,0,0,0])
                  PSE_T := pose_RPY2RotVec(p[0,0,0.005,0,0,0])
                  PSE_T_H := pose_trans(PSE_T, p[0,0,-0.008,0,0,0])
                  PSE_A := pose_trans(PSE_T, p[0,0,0.1,0,0,0])
                  PSE_R := pose_add(PSE_T, p[0,0,0.100,0,0,0])
            Case (caseValue=7)
              Folder define poses Manual
                GRP_Open_Pos := 60
                FRM_Reference := uLM_Manual
                If Action≟1
                  SuppressedNode
                    PSE_T := pose_RPY2RotVec(p[0.0202*(JIG_Slot%10),0.0202*(floor(JIG_Slot/10)),0,0,0,0])
                  PSE_T := pose_RPY2RotVec(p[0.0248*(JIG_Slot%8),0.0258*(floor(JIG_Slot/8)),0,0,0,0])
                  PSE_R := pose_add(PSE_T, p[0,0,0.150,0,0,0])
                ElseIf Action≟2
                  SuppressedNode
                    PSE_T := pose_RPY2RotVec(p[0.0202*(JIG_Slot%10),0.0202*(floor(JIG_Slot/10)),0,0,0,-62])
                  PSE_T := pose_RPY2RotVec(p[0.0248*(JIG_Slot%8),0.0258*(floor(JIG_Slot/8)),0,0,0,0])
                  PSE_R := pose_add(PSE_T, p[0,0,0.100,0,0,0])
                Script: PSE_T[2]=PSE_T[2]+PRM_TubHghtDiff
                PSE_A := pose_add(PSE_T, p[0,0,0.1,0,0,0])
      Case (caseValue=2)
        Folder Biorad
          'CHANGE THE REFERENCE TO THE FRAME TO MOVE IN'
          Folder Gripping parameters [hidden by the author, left out]
          If PRC_Target≟0
            Script: FRM_Reference = uML_BradRacks
            PSE_T := pose_RPY2RotVec(p[0.04365*JIG_Slot,0,0,0,0,180])
            If Action≟2
              SuppressedNode
                Script: PSE_T[2]=PSE_T[2]+0.008
              Script: PSE_T[2]=PSE_T[2]+0.002
            PSE_A := pose_add(PSE_T, p[0,0,0.18,0,0,0])
            PSE_R := pose_add(PSE_T, p[0,0,0.18,0,0,0])
          Else 
            Script: FRM_Reference = FRM_BioradMachn
            Switch expression=Action
              Case (caseValue=1)
                PSE_T := pose_RPY2RotVec(p[0.125-0.056*JIG_Slot,0.07,0.139,-90,0,0])
                PSE_A := pose_add(PSE_T, p[0,0.1,0,0,0,0])
                PSE_R := pose_add(PSE_T, p[0,0.05,0.1,0,0,0])
              Case (caseValue=2)
                PSE_T := pose_RPY2RotVec(p[0.125-0.056*JIG_Slot,0.07,0.08,-90,0,0])
                PSE_T_H := pose_RPY2RotVec(p[0.125-0.056*JIG_Slot,0.072,0.238,-90,0,0])
                PSE_A := pose_add(PSE_T_H, p[0,0.1,0,0,0,0])
                PSE_R := pose_add(PSE_T_H, p[0,0.1,0,0,0,0])
              Case (caseValue=7)
                PSE_T := pose_RPY2RotVec(p[0.124-0.056*JIG_Slot,0.084,0.008,-55,0,0])
                PSE_T_H := pose_RPY2RotVec(p[0.125-0.056*JIG_Slot,0.084,0.284,-55,0,0])
                PSE_A := pose_add(PSE_T_H, p[0,0.05,0.05,0,0,0])
                PSE_R := pose_add(PSE_T, p[0,0,0.1,0,0,0])
                SuppressedNode
                  JNT_Q := [0.108,-1.505,-1.993,-0.886,1.488,3.189]
              Case (caseValue=8)
                PSE_T_H := pose_RPY2RotVec(p[0.124-0.056*JIG_Slot,0.092,0.049,-72,0,0])
                PSE_T := pose_RPY2RotVec(p[0.125-0.056*JIG_Slot,0.092,0.316,-72,0,0])
                PSE_R := pose_add(PSE_T, p[0,0.05,0,0,0,0])
                PSE_A := pose_add(PSE_T_H, p[0,0,0.1,0,0,0])
                JNT_Q := [0.108,-1.505,-1.993,-0.886,1.488,3.189]
                If JIG_Slot≟0
                  Script: PSE_T[0]=PSE_T[0]-0.002
                  Script: PSE_T_H[0]=PSE_T_H[0]-0.002
      Case (caseValue=4)
        Folder Centrifuge
          'CHANGE THE REFERENCE TO THE FRAME TO MOVE IN'
          Folder Gripping parameters [hidden by the author, left out]
          If PRC_Target≟0
            Script: FRM_Reference = uLM_CentRacks
            Switch expression=Action
              Case (caseValue=1)
                PSE_T := pose_RPY2RotVec(p[0.0975*(JIG_Slot%4),0,-0.015,0,0,0])
              Case (caseValue=2)
                PSE_T := pose_RPY2RotVec(p[0.0975*(JIG_Slot%4),0,0.01,0,0,0])
            PSE_A := pose_add(PSE_T, p[0,0,0.15,0,0,0])
            PSE_R := pose_add(PSE_T, p[0,0,0.15,0,0,0])
          Else 
            Script: FRM_Reference = FRM_Centrifuge
            Switch expression=Action
              Case (caseValue=1)
                PSE_T := pose_RPY2RotVec(p[0,0,-0.02,0,0,0])
              Case (caseValue=2)
                PSE_T := pose_RPY2RotVec(p[0,0,0.015,0,0,0])
            PSE_A := pose_add(PSE_T, p[0,0,0.2,0,0,0])
            PSE_R := pose_add(PSE_T, p[0,0,0.25,0,0,0])
    Folder Additional check
      If not is_reachable(FRM_Reference,[PSE_A,PSE_A_H,PSE_T,PSE_T_H,PSE_R,PSE_R_H])
        Script: set_error(1002)
        Action := 0
  Switch expression=Action
    Case (caseValue=1)
      Folder Pick
        Action_Info := "Pick Rack/Probe"
        Script: do_transition(pose_trans(FRM_Reference, PSE_T), keep_rxry=OBJ_Picked)
        If not OBJ_Picked
          Script: rq_move_and_wait_norm(GRP_Open_Pos)
        If JNT_Q≠JNT_Z
          Script: movej(get_inverse_kin(pose_trans(FRM_Reference, PSE_A), qnear=JNT_Q))
        Else 
          MoveJ speed 100 deg/s, acceleration 80 deg/s^2 (useActiveTCP=true) feature=FRM_Reference
            Waypoint Variable (Variable): variable=PSE_A
        If ITM_ID≟4 and PRC_Target≟1
          Script: execute_cent_action(eACT_Inspect,(JIG_Slot+1))
        MoveL speed 400 mm/s, acceleration 500 mm/s^2 (useActiveTCP=true) feature=FRM_Reference
          Waypoint Variable (Variable): motionParameters(jointSpeed=1.047198 jointAcceleration=1.396263 cartesianSpeed=0.12 cartesianAcceleration=0.08); variable=PSE_T
          Script: rq_set_force_norm(50)
          SuppressedNode
            Script: rq_move_and_wait_norm(GRP_Close_Pos)
          URCap Gripper (Robotiq_Grippers, Robotiq Inc.) dataModel(position=100.0, force=76.0, speed=100.0, positionInDouble=100.0, forceInDouble=76.0, speedInDouble=100.0, slaveIds=[9], blocking=true)
          OBJ_Picked := rq_is_object_detected()
          Script: textmsg("Obj_Picked=",OBJ_Picked)
          If OBJ_Picked
            If PSE_T_H≠PSE_Z
              Waypoint Variable (Variable): motionParameters(blendRadius=0.01); variable=PSE_T_H
            Waypoint Variable (Variable): variable=PSE_R
          Else 
            Script: set_error(1010)
    Case (caseValue=2)
      Folder Place
        Action_Info := "place object"
        SuppressedNode
          Script: do_transition(keep_rxry=OBJ_Picked)
        Script: do_transition(pose_trans(FRM_Reference, PSE_T), keep_rxry=OBJ_Picked)
        If JNT_A≠[0,0,0,0,0,0]
          MoveJ speed 100 deg/s, acceleration 80 deg/s^2 (useActiveTCP=true positionType=JointAngles) feature=FRM_Reference
            Waypoint Variable (Variable): motionParameters(blendRadius=0.02); variable=JNT_A
        Else 
          MoveJ speed 100 deg/s, acceleration 80 deg/s^2 (useActiveTCP=true) feature=FRM_Reference
            Waypoint Variable (Variable): variable=PSE_A
        MoveL speed 400 mm/s, acceleration 500 mm/s^2 (useActiveTCP=true) feature=FRM_Reference
          If PSE_T_H≠PSE_Z
            Waypoint Variable (Variable): motionParameters(jointSpeed=1.047198 jointAcceleration=1.396263 cartesianSpeed=0.07 cartesianAcceleration=0.04); variable=PSE_T_H
          If ITM_ID≟4 and PRC_Target≟1
            Script: execute_cent_action(eACT_Inspect,(JIG_Slot+1))
          If not ERROR.FLAG
            If (ITM_ID≟1 and (JIG≟4 or JIG≟2)) or ITM_ID≟2 or ITM_ID≟4
              Waypoint Variable (Variable): motionParameters(jointSpeed=1.047198 jointAcceleration=1.396263 cartesianSpeed=0.09 cartesianAcceleration=0.05); variable=PSE_T
            Else 
              Waypoint Variable (Variable): motionParameters(jointSpeed=1.047198 jointAcceleration=1.396263 cartesianSpeed=0.09 cartesianAcceleration=0.05); variable=PSE_T
                Until TOOL_CONTACT_DETECTION (allowActions=false retraction=0 decelerationAcceleration=0.5 decelerationAngularAcceleration=34.906585)
              Force Frame feature=FRM_Reference; selection=[1, 1, 0, 0, 0, 0]; wrench=[0, 0, 0, 0, 0, 0]; limitsForce=[0.05, 0.05, 0.15, 1.047198, 1.047198, 1.047198]; limitsMotion=[0.1, 0.1, 0.1, 0.349066, 0.349066, 0.349066]
                Waypoint Variable (Variable): motionParameters(jointSpeed=1.047198 jointAcceleration=1.396263 cartesianSpeed=0.07 cartesianAcceleration=0.04); variable=PSE_T
            Script: rq_move_and_wait_norm(GRP_Open_Pos)
            Wait Sleep waitTime=0.2
            Waypoint Variable (Variable): variable=PSE_R
        SuppressedNode
          PRC_Task_Boxes := PRC_Task_Boxes+GRP_Boxes_Numb
    Case (caseValue=3)
      Folder Pick decapped probe from 3finger
        Action_Info := "Pick Rack/Probe"
        MoveJ speed 100 deg/s, acceleration 80 deg/s^2 (useActiveTCP=true) feature=FRM_Reference
          Waypoint Variable (Variable): variable=PSE_A
        Script: rq_move_and_wait_norm(GRP_Open_Pos)
        MoveL speed 75 mm/s, acceleration 150 mm/s^2 (useActiveTCP=true) feature=FRM_Reference
          SuppressedNode
            Script: PSE_T[2]=PSE_T[2]-0.005
          Waypoint Variable (Variable): variable=PSE_T
          SuppressedNode
            Force Frame feature=FRM_Reference; selection=[1, 1, 0, 0, 0, 0]; wrench=[0, 0, 0, 0, 0, 0]; limitsForce=[0.25, 0.25, 0.15, 1.047198, 1.047198, 1.047198]; limitsMotion=[0.1, 0.1, 0.1, 0.349066, 0.349066, 0.349066]
              Waypoint Variable (Variable): motionParameters(jointSpeed=1.047198 jointAcceleration=1.396263 cartesianSpeed=0.03 cartesianAcceleration=0.2); variable=PSE_T
          'ADD OPEN GRIPPER'
          Script: rq_set_force_norm(20)
          Script: rq_set_speed_norm(30)
          Script: rq_move_and_wait_norm(GRP_Close_Pos)
        Set DigitalOutput pin=digital_out[4]; digitalValue=1
        Wait Sleep waitTime=0.3
        MoveL speed 100 mm/s, acceleration 1200 mm/s^2 (useActiveTCP=true) feature=FRM_Reference
          Waypoint Variable (Variable): motionParameters(jointSpeed=1.047198 jointAcceleration=1.396263 cartesianSpeed=0.25 cartesianAcceleration=1.2); variable=PSE_R
    Case (caseValue=4)
      Folder Place probe in 3finger
        Action_Info := "place object"
        MoveJ speed 100 deg/s, acceleration 80 deg/s^2 (useActiveTCP=true) feature=FRM_Reference
          Waypoint Variable (Variable): variable=PSE_A
        Set DigitalOutput pin=digital_out[4]; digitalValue=1
        MoveL speed 75 mm/s, acceleration 150 mm/s^2 (useActiveTCP=true) feature=FRM_Reference
          Waypoint Variable (Variable): variable=PSE_T
            Until TOOL_CONTACT_DETECTION (allowActions=false retraction=0 decelerationAcceleration=3 decelerationAngularAcceleration=34.906585)
        Set DigitalOutput pin=digital_out[4]; digitalValue=0
        Wait Sleep waitTime=0.5
        SuppressedNode
          If Task_ID≟12
            Wait Sleep waitTime=0.15
            MoveL speed 75 mm/s, acceleration 150 mm/s^2 (useActiveTCP=true) feature=FRM_Reference
              Waypoint Variable (Variable): variable=PSE_R
    Case (caseValue=5)
      SuppressedNode
        Folder Decapping
          Action_Info := "decapping"
          PRM_decap_Zval := z_Pos
          PRM_forcdistSta := 0.02
          Script: zero_ftsensor()
          Wait Sleep waitTime=1
          Set DigitalOutput pin=digital_out[5]; digitalValue=1
          Set DigitalOutput pin=digital_out[3]; digitalValue=1
          Force Frame feature=uML_3fingergrip; selection=[0, 0, 1, 0, 0, 0]; wrench=[0, 0, 5, 0, 0, 0]; limitsForce=[0.04, 0.04, 0.015, 1.047198, 1.047198, 1.047198]; limitsMotion=[0.1, 0.1, 0.1, 0.349066, 0.349066, 0.349066]
            PRC_Force_Decap := True
            Wait Condition expression=PRM_forcdistLiv>PRM_forcdistSta
          PRC_Force_Decap := False
          Set DigitalOutput pin=digital_out[5]; digitalValue=0
          Set DigitalOutput pin=digital_out[3]; digitalValue=0
          MoveL speed 150 mm/s, acceleration 800 mm/s^2 (useActiveTCP=true) feature=FRM_Reference
            Waypoint Variable (Variable): variable=PSE_R
      Folder Decapping
        Action_Info := "decapping"
        Set DigitalOutput pin=digital_out[5]; digitalValue=1
        Set DigitalOutput pin=digital_out[3]; digitalValue=1
        Script: action_manipulator_decapping()
        Set DigitalOutput pin=digital_out[5]; digitalValue=0
        Set DigitalOutput pin=digital_out[3]; digitalValue=0
        MoveL speed 150 mm/s, acceleration 800 mm/s^2 (useActiveTCP=true) feature=FRM_Reference
          Waypoint Variable (Variable): variable=PSE_R
    Case (caseValue=6)
      SuppressedNode
        Folder Drop the cap
          Script: rq_set_speed_norm(100)
          Script: rq_set_force_norm(10)
          MoveJ speed 100 deg/s, acceleration 80 deg/s^2 (useActiveTCP=true) feature=FRM_Reference
            Waypoint Variable (Variable): motionParameters(blendRadius=0.02); variable=PSE_A
          MoveL speed 400 mm/s, acceleration 500 mm/s^2 (useActiveTCP=true) feature=FRM_Reference
            Waypoint Variable (Variable): motionParameters(jointSpeed=1.047198 jointAcceleration=1.396263 cartesianSpeed=0.09 cartesianAcceleration=0.05); variable=PSE_T
            'ADD OPEN GRIPPER'
            Loop While (checkContinuously=false) expression=rq_is_object_detected()
              URCap Gripper (Robotiq_Grippers, Robotiq Inc.) dataModel(position=0.0, force=28.0, speed=100.0, positionInDouble=0.0, forceInDouble=28.0, speedInDouble=100.0, slaveIds=[9], blocking=true)
              Wait Sleep waitTime=0.01
              URCap Gripper (Robotiq_Grippers, Robotiq Inc.) dataModel(position=100.0, force=28.0, speed=100.0, positionInDouble=100.0, forceInDouble=28.0, speedInDouble=100.0, slaveIds=[9], blocking=true)
            Wait Sleep waitTime=0.2
            Waypoint Variable (Variable): variable=PSE_R
      Folder Drop
        Script: rq_set_speed_norm(100)
        MoveJ speed 100 deg/s, acceleration 80 deg/s^2 (useActiveTCP=true) feature=FRM_Reference
          Waypoint Variable (Variable): motionParameters(blendRadius=0.02); variable=PSE_A
        MoveL speed 400 mm/s, acceleration 500 mm/s^2 (useActiveTCP=true) feature=FRM_Reference
          Waypoint Variable (Variable): motionParameters(jointSpeed=1.047198 jointAcceleration=1.396263 cartesianSpeed=0.12 cartesianAcceleration=0.08); variable=PSE_T
          URCap Gripper (Robotiq_Grippers, Robotiq Inc.) dataModel(position=70.19607843137254, force=30.19607843137255, speed=0.0, positionInDouble=70.19607843137254, forceInDouble=30.19607843137255, speedInDouble=0.0, slaveIds=[9], blocking=true)
          Waypoint Variable (Variable): motionParameters(jointSpeed=1.047198 jointAcceleration=1.396263 cartesianSpeed=0.12 cartesianAcceleration=0.08); variable=PSE_T_H
          Script: rq_move_and_wait_norm(GRP_Open_Pos)
          Wait Sleep waitTime=0.2
          Waypoint Variable (Variable): variable=PSE_R
    Case (caseValue=7)
      Folder Load
        Action_Info := "load object in the machine"
        SuppressedNode
          Script: do_transition(keep_rxry=OBJ_Picked)
        If JNT_Q≠JNT_Z
          Script: movej(get_inverse_kin(pose_trans(FRM_Reference, PSE_A), qnear=JNT_Q), r=0.05)
        Else 
          MoveJ speed 100 deg/s, acceleration 80 deg/s^2 (useActiveTCP=true) feature=FRM_Reference
            Waypoint Variable (Variable): motionParameters(blendRadius=0.02); variable=PSE_A
        MoveL speed 400 mm/s, acceleration 500 mm/s^2 (useActiveTCP=true) feature=FRM_Reference
          SuppressedNode
            Waypoint Variable (Variable): motionParameters(jointSpeed=1.047198 jointAcceleration=1.396263 cartesianSpeed=0.09 cartesianAcceleration=0.05); variable=PSE_T
              Until TOOL_CONTACT_DETECTION (allowActions=false retraction=0 decelerationAcceleration=0.5 decelerationAngularAcceleration=34.906585)
          SuppressedNode
            Force Frame feature=FRM_Reference; selection=[1, 1, 0, 0, 0, 0]; wrench=[0, 0, 0, 0, 0, 0]; limitsForce=[0.05, 0.05, 0.15, 1.047198, 1.047198, 1.047198]; limitsMotion=[0.1, 0.1, 0.1, 0.349066, 0.349066, 0.349066]
              Waypoint Variable (Variable): motionParameters(jointSpeed=1.047198 jointAcceleration=1.396263 cartesianSpeed=0.07 cartesianAcceleration=0.04); variable=PSE_T
          Waypoint Variable (Variable): motionParameters(jointSpeed=1.047198 jointAcceleration=1.396263 cartesianSpeed=0.07 cartesianAcceleration=0.04); variable=PSE_T_H
          URCap Gripper (Robotiq_Grippers, Robotiq Inc.) dataModel(position=100.0, force=0.0, speed=67.84313725490196, positionInDouble=100.0, forceInDouble=0.0, speedInDouble=67.84313725490196, slaveIds=[9], blocking=true)
          Wait Sleep waitTime=0.2
          Waypoint Variable (Variable): motionParameters(jointSpeed=1.047198 jointAcceleration=1.396263 cartesianSpeed=0.07 cartesianAcceleration=0.04); variable=PSE_T
          Waypoint Variable (Variable): variable=PSE_R
    Case (caseValue=8)
      Folder UnLoad
        Action_Info := "unload object in the machine"
        SuppressedNode
          Script: do_transition(keep_rxry=OBJ_Picked)
        If JNT_Q≠JNT_Z
          SuppressedNode
            Script: movej(get_inverse_kin(pose_trans(FRM_Reference, PSE_A), qnear=JNT_Q), r=0.01)
          Script: movej(get_inverse_kin(pose_trans(FRM_Reference, PSE_A), qnear=JNT_Q))
        Else 
          MoveJ speed 100 deg/s, acceleration 80 deg/s^2 (useActiveTCP=true) feature=FRM_Reference
            Waypoint Variable (Variable): variable=PSE_A
        MoveL speed 400 mm/s, acceleration 500 mm/s^2 (useActiveTCP=true) feature=FRM_Reference
          SuppressedNode
            Waypoint Variable (Variable): motionParameters(jointSpeed=1.047198 jointAcceleration=1.396263 cartesianSpeed=0.09 cartesianAcceleration=0.05); variable=PSE_T
              Until TOOL_CONTACT_DETECTION (allowActions=false retraction=0 decelerationAcceleration=0.5 decelerationAngularAcceleration=34.906585)
          SuppressedNode
            Force Frame feature=FRM_Reference; selection=[1, 1, 0, 0, 0, 0]; wrench=[0, 0, 0, 0, 0, 0]; limitsForce=[0.05, 0.05, 0.15, 1.047198, 1.047198, 1.047198]; limitsMotion=[0.1, 0.1, 0.1, 0.349066, 0.349066, 0.349066]
              Waypoint Variable (Variable): motionParameters(jointSpeed=1.047198 jointAcceleration=1.396263 cartesianSpeed=0.07 cartesianAcceleration=0.04); variable=PSE_T
          Script: rq_move_and_wait_norm(GRP_Open_Pos)
          Waypoint Variable (Variable): motionParameters(jointSpeed=1.047198 jointAcceleration=1.396263 cartesianSpeed=0.07 cartesianAcceleration=0.04); variable=PSE_T_H
          URCap Gripper (Robotiq_Grippers, Robotiq Inc.) dataModel(position=100.0, force=0.0, speed=67.84313725490196, positionInDouble=100.0, forceInDouble=0.0, speedInDouble=67.84313725490196, slaveIds=[9], blocking=true)
          Wait Sleep waitTime=0.2
          OBJ_Picked := rq_is_object_detected()
          If OBJ_Picked
            Waypoint Variable (Variable): motionParameters(jointSpeed=1.047198 jointAcceleration=1.396263 cartesianSpeed=0.07 cartesianAcceleration=0.04); variable=PSE_T
            Script: rq_move_and_wait_norm(GRP_Open_Pos)
            Waypoint Variable (Variable): variable=PSE_R
          Else 
            Script: set_error(1010)
    Case (caseValue=16)
      Folder Scan the barcode
        Action_Info := "scan the barcode"
        Barc_scan_succs := False
        Folder First check
          Set DigitalOutput pin=digital_out[6]; digitalValue=1
          Wait Sleep waitTime=0.1
          Barc_scan_succs := digital_in[6]
        If Barc_scan_succs
          Set DigitalOutput pin=digital_out[5]; digitalValue=1
          Set DigitalOutput pin=digital_out[2]; digitalValue=1
          Loop While (checkContinuously=true) expression=Barc_scan_succs
            Barc_scan_succs := digital_in[6]
            Wait Sleep waitTime=0.05
          Set DigitalOutput pin=digital_out[5]; digitalValue=0
          Set DigitalOutput pin=digital_out[2]; digitalValue=0
          Set DigitalOutput pin=digital_out[6]; digitalValue=0
        Else 
          Timer (action=Reset) variable(name=Timer_Barc_scan)
          Timer (action=Start) variable=Timer_Barc_scan
          Set DigitalOutput pin=digital_out[3]; digitalValue=1
          Set DigitalOutput pin=digital_out[5]; digitalValue=1
          Loop While (checkContinuously=true) expression=not Barc_scan_succs and  not CMD_Stop and Timer_Barc_scan<60
            SuppressedNode
              If Timer_Barc_scan>1.5
                Placeholder
            Set DigitalOutput pin=digital_out[6]; digitalValue=1
            Barc_scan_succs := digital_in[6]
            Wait Sleep waitTime=0.05
          Set DigitalOutput pin=digital_out[5]; digitalValue=0
          Set DigitalOutput pin=digital_out[3]; digitalValue=0
          Set DigitalOutput pin=digital_out[6]; digitalValue=0
          Timer (action=Stop) variable=Timer_Barc_scan
          If Timer_Barc_scan≥60
            Script: set_error(5200)
  '=========='
  Script: textmsg("Action=",Action)
  Folder PostSettings [hidden by the author, left out]
